// TIA Portal V21 export
// export: Created 2026-11-18T10:00:00.0000000Z, ExportSetting None
FUNCTION_BLOCK "FB_Station"   // FB20, LAD
{ S7_Optimized_Access := 'TRUE' }
// stored: MemoryReserve 100, SetENOAutomatically false
   VAR_INPUT
      Enable : Bool;
      Init : Bool;
   END_VAR
   VAR_OUTPUT
      Lamp : Bool;
   END_VAR
   VAR
      Seq : "FB_Sequence";
      Run : Bool;
   END_VAR
BEGIN

REGION Network 1: Sequence
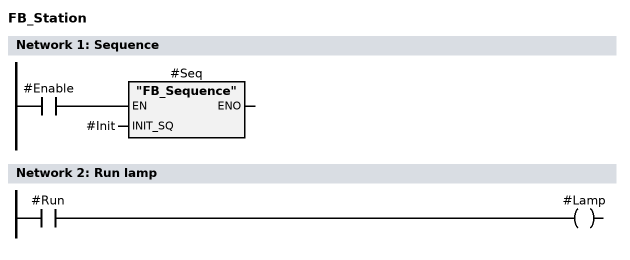
   RUNG wire#powerrail
      Contact( #Enable )
      #Seq(INIT_SQ := #Init)
   END_RUNG
   // the same network as SCL:
   IF #Enable THEN
       #Seq(INIT_SQ := #Init);   // "FB_Sequence"
   END_IF;
END_REGION

REGION Network 2: Run lamp
   RUNG wire#powerrail
      Contact( #Run )
      Coil( #Lamp )
   END_RUNG
   // the same network as SCL:
   #Lamp := #Run;
END_REGION
END_FUNCTION_BLOCK
